// TIA Portal V20 export
FUNCTION_BLOCK "FB_LD_PressDemoLoadPosition"   // FB, LAD
{ S7_Optimized_Access := 'TRUE' }
// stored: AutoNumber true
   VAR_INPUT
      Run { ExternalWritable := 'False'} : Bool;
      Reset { ExternalWritable := 'False'} : Bool;
      OwnerIndex { ExternalWritable := 'False'} : DInt;
      Delta { ExternalWritable := 'False'} : Time;
   END_VAR
   VAR_IN_OUT
      PressRam { ExternalAccessible := 'False'; ExternalVisible := 'False'; ExternalWritable := 'False'} : "FB_CylinderCM";
      Door { ExternalAccessible := 'False'; ExternalVisible := 'False'; ExternalWritable := 'False'} : "FB_CylinderCM";
      PartSlide { ExternalAccessible := 'False'; ExternalVisible := 'False'; ExternalWritable := 'False'} : "FB_CylinderCM";
   END_VAR
   VAR
      Seq { ExternalWritable := 'False'} : "FRK_SequenceCtx";
      Row1 { ExternalWritable := 'False'} : "FRK_SequenceRow";
      Row2 { ExternalWritable := 'False'} : "FRK_SequenceRow";
      Row3 { ExternalWritable := 'False'} : "FRK_SequenceRow";
      Row4 { ExternalWritable := 'False'} : "FRK_SequenceRow";
      At240 { ExternalAccessible := 'False'; ExternalVisible := 'False'; ExternalWritable := 'False'} : Bool;
      At260 { ExternalAccessible := 'False'; ExternalVisible := 'False'; ExternalWritable := 'False'} : Bool;
      At280 { ExternalAccessible := 'False'; ExternalVisible := 'False'; ExternalWritable := 'False'} : Bool;
      At300 { ExternalAccessible := 'False'; ExternalVisible := 'False'; ExternalWritable := 'False'} : Bool;
      Ready1 { ExternalAccessible := 'False'; ExternalVisible := 'False'; ExternalWritable := 'False'} : Bool;
      Ready2 { ExternalAccessible := 'False'; ExternalVisible := 'False'; ExternalWritable := 'False'} : Bool;
      Ready3 { ExternalAccessible := 'False'; ExternalVisible := 'False'; ExternalWritable := 'False'} : Bool;
      Ready4 { ExternalAccessible := 'False'; ExternalVisible := 'False'; ExternalWritable := 'False'} : Bool;
      Ready5 { ExternalAccessible := 'False'; ExternalVisible := 'False'; ExternalWritable := 'False'} : Bool;
      Advance { ExternalAccessible := 'False'; ExternalVisible := 'False'; ExternalWritable := 'False'} : Bool;
   END_VAR
BEGIN

REGION Network 1
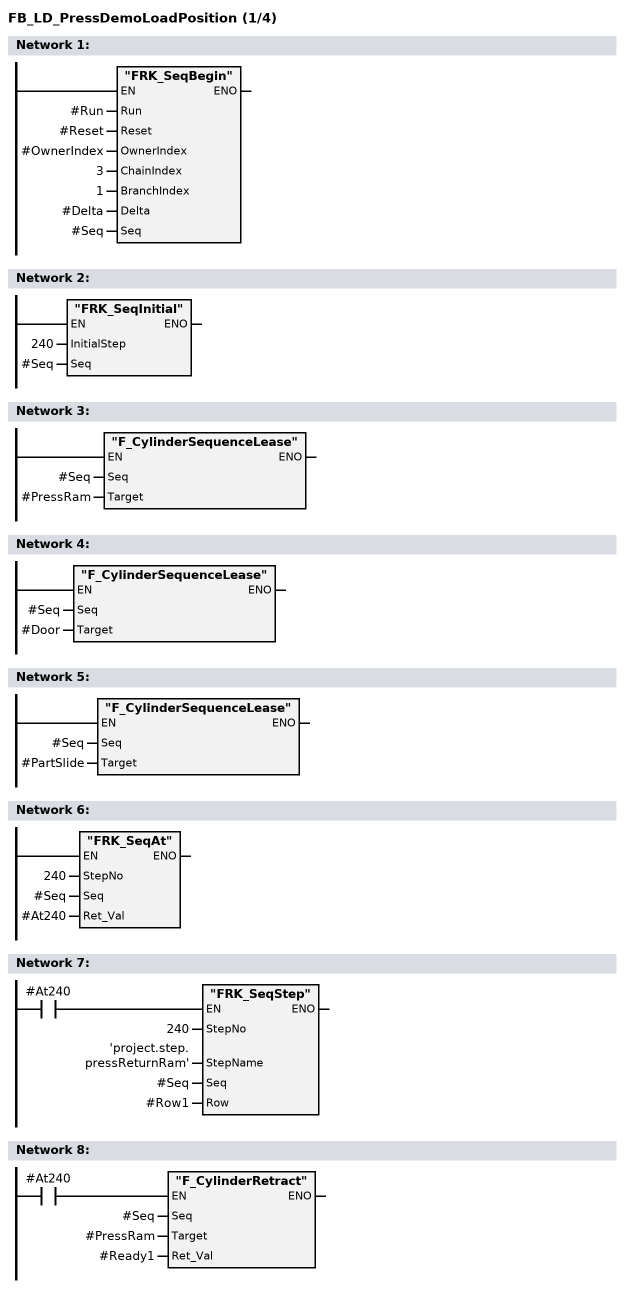
   RUNG wire#powerrail
      "FRK_SeqBegin"(Run := #Run, Reset := #Reset, OwnerIndex := #OwnerIndex, ChainIndex := 3, BranchIndex := 1, Delta := #Delta, Seq := #Seq)
   END_RUNG
   // the same network as SCL:
   "FRK_SeqBegin"(Run := #Run,
                  Reset := #Reset,
                  OwnerIndex := #OwnerIndex,
                  ChainIndex := 3,
                  BranchIndex := 1,
                  Delta := #Delta,
                  Seq := #Seq);
END_REGION

REGION Network 2
   RUNG wire#powerrail
      "FRK_SeqInitial"(InitialStep := 240, Seq := #Seq)
   END_RUNG
   // the same network as SCL:
   "FRK_SeqInitial"(InitialStep := 240, Seq := #Seq);
END_REGION

REGION Network 3
   RUNG wire#powerrail
      "F_CylinderSequenceLease"(Seq := #Seq, Target := #PressRam)
   END_RUNG
   // the same network as SCL:
   "F_CylinderSequenceLease"(Seq := #Seq, Target := #PressRam);
END_REGION

REGION Network 4
   RUNG wire#powerrail
      "F_CylinderSequenceLease"(Seq := #Seq, Target := #Door)
   END_RUNG
   // the same network as SCL:
   "F_CylinderSequenceLease"(Seq := #Seq, Target := #Door);
END_REGION

REGION Network 5
   RUNG wire#powerrail
      "F_CylinderSequenceLease"(Seq := #Seq, Target := #PartSlide)
   END_RUNG
   // the same network as SCL:
   "F_CylinderSequenceLease"(Seq := #Seq, Target := #PartSlide);
END_REGION

REGION Network 6
   RUNG wire#powerrail
      "FRK_SeqAt"(StepNo := 240, Seq := #Seq, Ret_Val := #At240)
   END_RUNG
   // the same network as SCL:
   "FRK_SeqAt"(StepNo := 240, Seq := #Seq, Ret_Val := #At240);
END_REGION

REGION Network 7
   IF #At240 THEN
       "FRK_SeqStep"(StepNo := 240, StepName := 'project.step.pressReturnRam', Seq := #Seq, Row := #Row1);
   END_IF;
END_REGION

REGION Network 8
   IF #At240 THEN "F_CylinderRetract"(Seq := #Seq, Target := #PressRam, Ret_Val := #Ready1); END_IF;
END_REGION

REGION Network 9
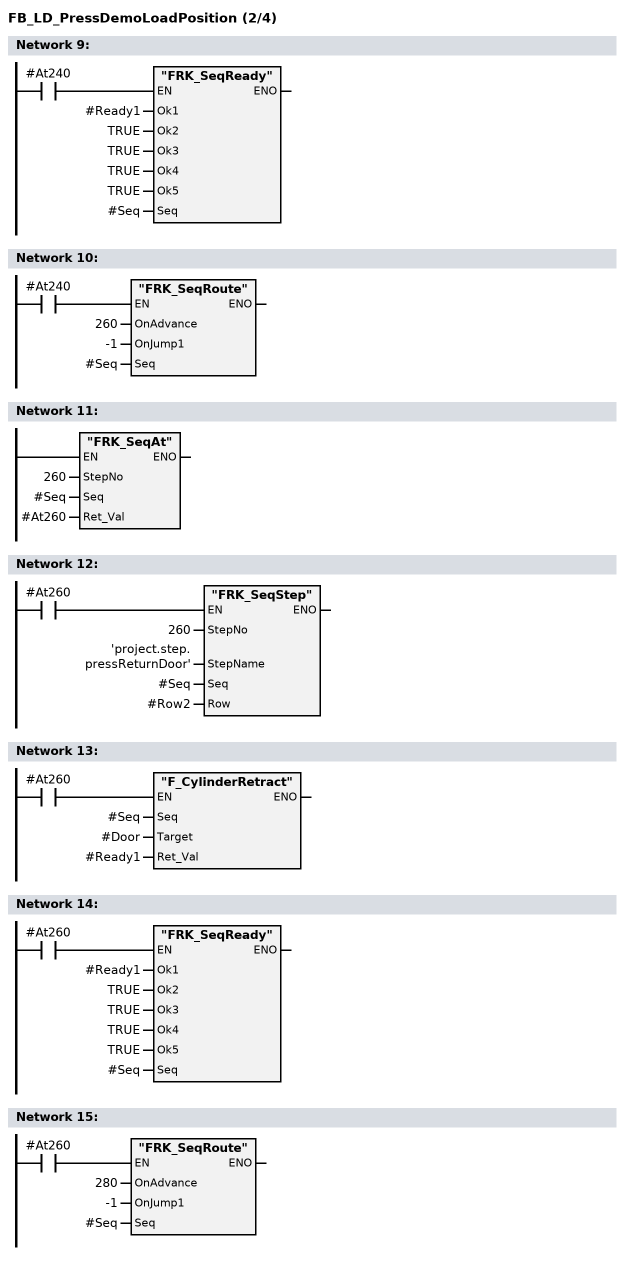
   IF #At240 THEN
       "FRK_SeqReady"(Ok1 := #Ready1, Ok2 := TRUE, Ok3 := TRUE, Ok4 := TRUE, Ok5 := TRUE, Seq := #Seq);
   END_IF;
END_REGION

REGION Network 10
   IF #At240 THEN "FRK_SeqRoute"(OnAdvance := 260, OnJump1 := -1, Seq := #Seq); END_IF;
END_REGION

REGION Network 11
   RUNG wire#powerrail
      "FRK_SeqAt"(StepNo := 260, Seq := #Seq, Ret_Val := #At260)
   END_RUNG
   // the same network as SCL:
   "FRK_SeqAt"(StepNo := 260, Seq := #Seq, Ret_Val := #At260);
END_REGION

REGION Network 12
   IF #At260 THEN
       "FRK_SeqStep"(StepNo := 260, StepName := 'project.step.pressReturnDoor', Seq := #Seq, Row := #Row2);
   END_IF;
END_REGION

REGION Network 13
   IF #At260 THEN "F_CylinderRetract"(Seq := #Seq, Target := #Door, Ret_Val := #Ready1); END_IF;
END_REGION

REGION Network 14
   IF #At260 THEN
       "FRK_SeqReady"(Ok1 := #Ready1, Ok2 := TRUE, Ok3 := TRUE, Ok4 := TRUE, Ok5 := TRUE, Seq := #Seq);
   END_IF;
END_REGION

REGION Network 15
   IF #At260 THEN "FRK_SeqRoute"(OnAdvance := 280, OnJump1 := -1, Seq := #Seq); END_IF;
END_REGION

REGION Network 16
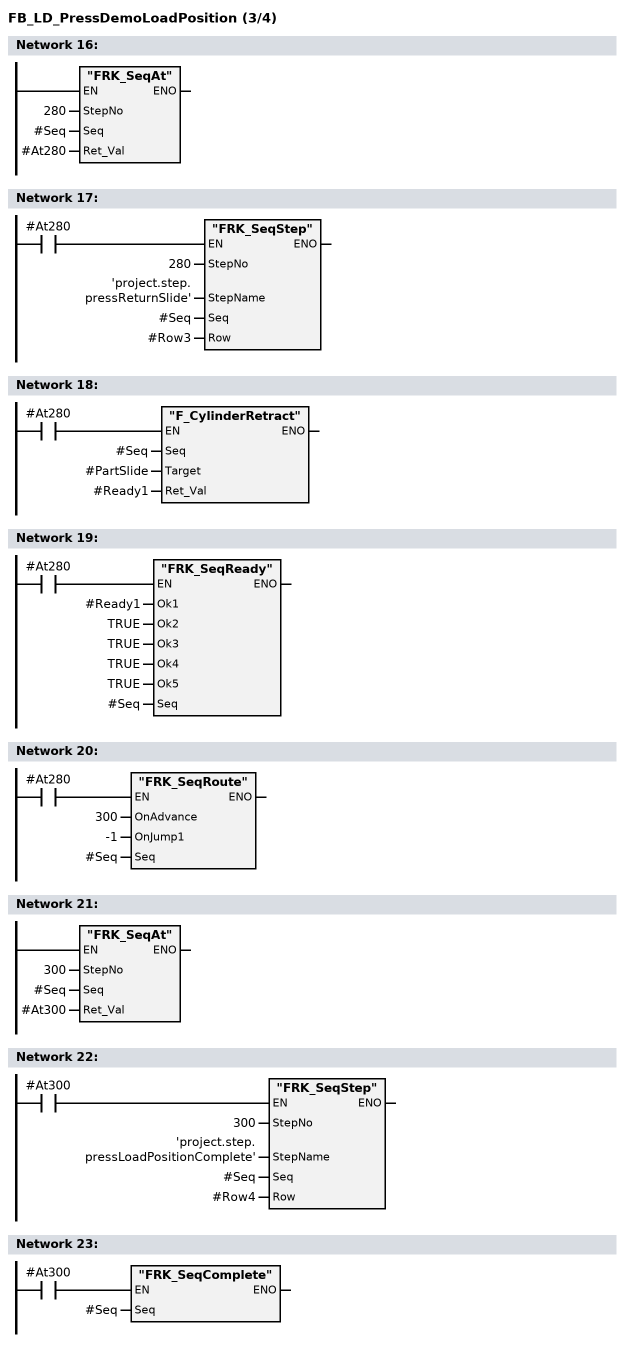
   RUNG wire#powerrail
      "FRK_SeqAt"(StepNo := 280, Seq := #Seq, Ret_Val := #At280)
   END_RUNG
   // the same network as SCL:
   "FRK_SeqAt"(StepNo := 280, Seq := #Seq, Ret_Val := #At280);
END_REGION

REGION Network 17
   IF #At280 THEN
       "FRK_SeqStep"(StepNo := 280, StepName := 'project.step.pressReturnSlide', Seq := #Seq, Row := #Row3);
   END_IF;
END_REGION

REGION Network 18
   IF #At280 THEN "F_CylinderRetract"(Seq := #Seq, Target := #PartSlide, Ret_Val := #Ready1); END_IF;
END_REGION

REGION Network 19
   IF #At280 THEN
       "FRK_SeqReady"(Ok1 := #Ready1, Ok2 := TRUE, Ok3 := TRUE, Ok4 := TRUE, Ok5 := TRUE, Seq := #Seq);
   END_IF;
END_REGION

REGION Network 20
   IF #At280 THEN "FRK_SeqRoute"(OnAdvance := 300, OnJump1 := -1, Seq := #Seq); END_IF;
END_REGION

REGION Network 21
   RUNG wire#powerrail
      "FRK_SeqAt"(StepNo := 300, Seq := #Seq, Ret_Val := #At300)
   END_RUNG
   // the same network as SCL:
   "FRK_SeqAt"(StepNo := 300, Seq := #Seq, Ret_Val := #At300);
END_REGION

REGION Network 22
   IF #At300 THEN
       "FRK_SeqStep"(StepNo := 300, StepName := 'project.step.pressLoadPositionComplete', Seq := #Seq, Row := #Row4);
   END_IF;
END_REGION

REGION Network 23
   IF #At300 THEN "FRK_SeqComplete"(Seq := #Seq); END_IF;
END_REGION

REGION Network 24
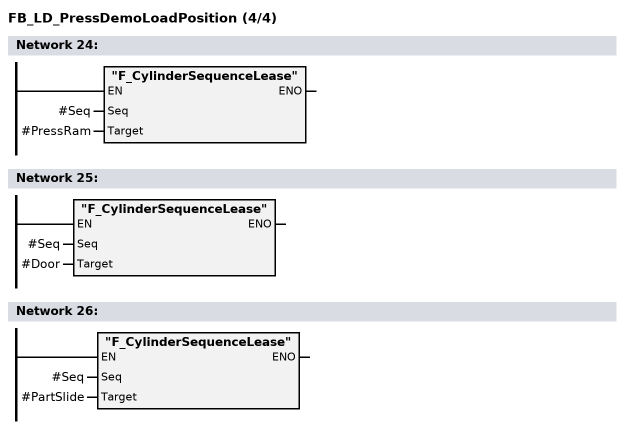
   RUNG wire#powerrail
      "F_CylinderSequenceLease"(Seq := #Seq, Target := #PressRam)
   END_RUNG
   // the same network as SCL:
   "F_CylinderSequenceLease"(Seq := #Seq, Target := #PressRam);
END_REGION

REGION Network 25
   RUNG wire#powerrail
      "F_CylinderSequenceLease"(Seq := #Seq, Target := #Door)
   END_RUNG
   // the same network as SCL:
   "F_CylinderSequenceLease"(Seq := #Seq, Target := #Door);
END_REGION

REGION Network 26
   RUNG wire#powerrail
      "F_CylinderSequenceLease"(Seq := #Seq, Target := #PartSlide)
   END_RUNG
   // the same network as SCL:
   "F_CylinderSequenceLease"(Seq := #Seq, Target := #PartSlide);
END_REGION
END_FUNCTION_BLOCK
